(* PLC project zarechnaya.project, CODESYS CODESYS V3.5 SP17 Patch 3 *)
(* stored: creationDateTime 2026-10-20T05:42:22.2150167, modificationDateTime 1601-01-01T03:00:00 *)

(* FB_ValveCmd — команда регулирующей задвижки (FBD, MOVE/SEL/LIMIT; EN/ENO не используется — M0: N). Поведение (модель scenarios/reference/model_FB_ValveCmd.py): 1. iCmd := SEL(xOpen, iClosedPos, iOpenPos) — xOpen = FALSE → iClosedPos, TRUE → iOpenPos; 2. iPos := LIMIT(iMin, iCmd, iMax); 3. iOut := MOVE(iPos); 4. xAtLimit := (iPos = iMin) OR (iPos = iMax). SEL и LIMIT вне подмножества FlgNet P0 → блок целиком в SCL (C2S7-GFX-SCL). *)
FUNCTION_BLOCK FB_ValveCmd
  VAR_INPUT
    xOpen : BOOL;
    iClosedPos : INT;
    iOpenPos : INT;
    iMin : INT;
    iMax : INT;
  END_VAR
  VAR_OUTPUT
    iOut : INT;
    xAtLimit : BOOL;
  END_VAR
  VAR
    iCmd : INT;
    iPos : INT;
  END_VAR

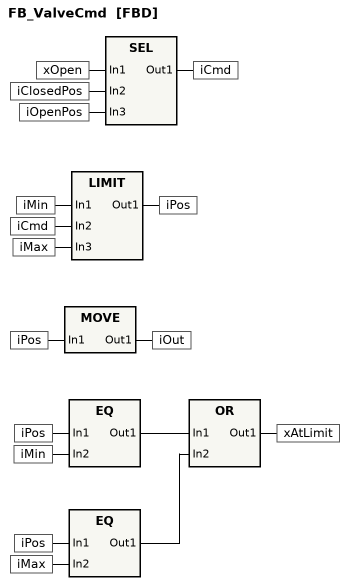
(* FBD diagram, written out as Structured Text *)
iCmd := SEL(xOpen, iClosedPos, iOpenPos);
(* --- network: Ограничение --- *)
iPos := LIMIT(iMin, iCmd, iMax);
(* --- network: Выход --- *)
iOut := iPos;
(* --- network: На упоре --- *)
xAtLimit := iPos = iMin OR iPos = iMax;
END_FUNCTION_BLOCK
